(* IEC 61131-3 sources: 2026_Projet_YGO_ExcavatriceDragage/TOOLS/TEST_AUTO_CI/RESULTS/L_SIMULATION/tests (part 4) *)

(* ---- test_fb_simbench.st ---- *)
SETUP
VAR
    FB_Bench : FB_SimBench;
    FB_SimEnc : FB_Sim_Encoder;
    FB_SimJoy : FB_Sim_Joystick;
    FB_SimSafe : FB_Sim_Safety;
    FB_SimTrans : FB_Sim_Translation;
    RawPosM1 : UDINT := 0;
    RawPosM2 : UDINT := 0;
END_VAR
END_SETUP

TEST 'TC-P03-001 Dynamique Enable : neutralisation initiale, transition Ready au repos, puis coupure'
    (* Scan 0 : Enable=FALSE -> Neutralisation *)
    FB_Bench(Enable := FALSE, RawPosM1 := RawPosM1, RawPosM2 := RawPosM2);
    ASSERT_FALSE(FB_Bench.Ready, 'Enable=FALSE -> Ready=FALSE (neutralise)');

    ADVANCE_TIME(10000000);

    (* Scan 1 : Enable=TRUE -> SimBench actif *)
    FB_Bench(Enable := TRUE, RawPosM1 := RawPosM1, RawPosM2 := RawPosM2);
    ASSERT_TRUE(FB_Bench.Ready, 'Enable=TRUE -> Ready=TRUE (nominal)');

    ADVANCE_TIME(10000000);

    (* Scan 2 : Enable=FALSE -> Re-neutralisation *)
    FB_Bench(Enable := FALSE, RawPosM1 := RawPosM1, RawPosM2 := RawPosM2);
    ASSERT_FALSE(FB_Bench.Ready, 'Coupure -> Ready retombe a FALSE');
END_TEST

(* =========================================================================
   T419 — Reprise de jeu : ne jamais ouvrir la benne pendant une descente M1+M2.
   ========================================================================= *)

TEST 'TC-P13-074 T419 descente M1-M2 : compensation de fermeture conservee'
VAR
    CorrectionAfterAscentPts       : DINT;
    CorrectionAfterBothDescentPts  : DINT;
END_VAR
    (* La montee couplee etablit une compensation de fermeture observable. *)
    RawPosM1 := 1000000; RawPosM2 := 1100000;
    FB_Bench(Enable := TRUE, RawPosM1 := RawPosM1, RawPosM2 := RawPosM2,
             M1_RelayFwd := TRUE, M2_RelayFwd := TRUE,
             M1_BrakeCmd := TRUE, M2_BrakeCmd := TRUE,
             SimWinchCouplingModelActive := TRUE,
             M1_CablePos_M := 5.0, M2_CablePos_M := 18.5,
             BucketOffsetCloseM := 15.0, BucketCoherenceLimitM := 1.0);
    ADVANCE_TIME(10000000);

    (* Second scan : reprise de jeu de fermeture accumulee dans l'image M2. *)
    FB_Bench(Enable := TRUE, RawPosM1 := RawPosM1, RawPosM2 := RawPosM2,
             M1_RelayFwd := TRUE, M2_RelayFwd := TRUE,
             M1_BrakeCmd := TRUE, M2_BrakeCmd := TRUE,
             SimWinchCouplingModelActive := TRUE,
             M1_CablePos_M := 5.0, M2_CablePos_M := 18.5,
             BucketOffsetCloseM := 15.0, BucketCoherenceLimitM := 1.0);
    CorrectionAfterAscentPts := UDINT_TO_DINT(FB_Bench.Winch.COD2_PosValue) - UDINT_TO_DINT(RawPosM2);
    ASSERT_TRUE(CorrectionAfterAscentPts > 0, 'montee couplee -> compensation fermee presente');
    ADVANCE_TIME(10000000);

    (* Descente de charge M1+M2 : ce n'est pas une ouverture relative de la benne. *)
    FB_Bench(Enable := TRUE, RawPosM1 := RawPosM1, RawPosM2 := RawPosM2,
             M1_RelayFwd := FALSE, M1_RelayRev := TRUE,
             M2_RelayFwd := FALSE, M2_RelayRev := TRUE,
             M1_BrakeCmd := TRUE, M2_BrakeCmd := TRUE,
             SimWinchCouplingModelActive := TRUE,
             M1_CablePos_M := 5.0, M2_CablePos_M := 18.5,
             BucketOffsetCloseM := 15.0, BucketCoherenceLimitM := 1.0);
    CorrectionAfterBothDescentPts := UDINT_TO_DINT(FB_Bench.Winch.COD2_PosValue) - UDINT_TO_DINT(RawPosM2);
    ASSERT_EQ(CorrectionAfterBothDescentPts, CorrectionAfterAscentPts,
              'descente M1+M2 -> compensation de fermeture inchangee');
END_TEST

TEST 'TC-P13-075 T419 ouverture M2 seule : relachement borne conserve'
VAR
    CorrectionBeforeOpenPts : DINT;
    CorrectionAfterOpenPts  : DINT;
END_VAR
    (* Scenario autonome : etabli une fermeture avant l'ouverture relative M2 seule. *)
    RawPosM1 := 1000000; RawPosM2 := 1100000;
    FB_Bench(Enable := TRUE, RawPosM1 := RawPosM1, RawPosM2 := RawPosM2,
             M1_RelayFwd := TRUE, M2_RelayFwd := TRUE,
             M1_BrakeCmd := TRUE, M2_BrakeCmd := TRUE,
             SimWinchCouplingModelActive := TRUE,
             M1_CablePos_M := 5.0, M2_CablePos_M := 18.5,
             BucketOffsetCloseM := 15.0, BucketCoherenceLimitM := 1.0);
    ADVANCE_TIME(10000000);
    CorrectionBeforeOpenPts := UDINT_TO_DINT(FB_Bench.Winch.COD2_PosValue) - UDINT_TO_DINT(RawPosM2);
    ASSERT_TRUE(CorrectionBeforeOpenPts > 0, 'fermeture etablie avant ouverture M2 seule');
    ADVANCE_TIME(10000000);
    FB_Bench(Enable := TRUE, RawPosM1 := RawPosM1, RawPosM2 := RawPosM2,
             M1_RelayFwd := FALSE, M1_RelayRev := FALSE,
             M2_RelayFwd := FALSE, M2_RelayRev := TRUE,
             M2_BrakeCmd := TRUE,
             SimWinchCouplingModelActive := TRUE,
             M1_CablePos_M := 5.0, M2_CablePos_M := 18.5,
             BucketOffsetCloseM := 15.0, BucketCoherenceLimitM := 1.0);
    CorrectionAfterOpenPts := UDINT_TO_DINT(FB_Bench.Winch.COD2_PosValue) - UDINT_TO_DINT(RawPosM2);
    ASSERT_TRUE(CorrectionAfterOpenPts < CorrectionBeforeOpenPts,
                'ouverture M2 seule -> compensation relachee');
    ASSERT_TRUE((CorrectionBeforeOpenPts - CorrectionAfterOpenPts) <= 82,
                'ouverture M2 seule -> relachement borne a 0,02 m par scan');
END_TEST

TEST 'TC-P13-001 Sim_Safety : neutralisation sans Enable'
    FB_SimSafe(Enable := FALSE);
    ASSERT_FALSE(FB_SimSafe.SimChainOk, 'AU non ferme');
    ASSERT_FALSE(FB_SimSafe.SimContactorOk, 'Contacteur coupe');
END_TEST

(* =========================================================================
   AF-13 — FB_SimBench (TC-P13-010/011/012/013)
   ========================================================================= *)

TEST 'TC-P13-010 SimBench Enable=FALSE neutralise tout le banc'
    FB_Bench(Enable := FALSE, RawPosM1 := RawPosM1, RawPosM2 := RawPosM2);
    ASSERT_FALSE(FB_Bench.Ready, 'Enable=FALSE -> Ready=FALSE');
    ASSERT_FALSE(FB_Bench.Busy, 'Enable=FALSE -> Busy=FALSE');
    ASSERT_FALSE(FB_Bench.Done, 'Enable=FALSE -> Done=FALSE');
END_TEST

(* =========================================================================
   T342 — CR2 : reinjection silencieuse du comptage brut (RawPosM2 = 0 -> 1 100 000 pts)
   Remplace TC-P13-014 « initialise les codeurs absolus vierges » (ID par ailleurs porte
   par l'AF-13 pour le capteur haut TOP : collision d'ID levee au passage) : le banc
   n'initialise PLUS rien, le cas « memoire vierge » est couvert par l'initialisation
   declaree GVL_PERSISTENT._SimEncoderRawPosM1/M2 := 1000000.
   ========================================================================= *)

TEST 'TC-T342-010 AUCUNE reinjection du comptage brut : un 0 reel du codeur est conserve (pas de saut post-AU)'
    (* Etat EXACT de l'incident T338 (saut 8,50 -> 204,677 m apres reactivation du banc) :
       memoire codeur a 0, banc desactive (Enable=FALSE), puis reactivation du banc
       (GVL_Simulation.SimulationModeActive FALSE -> TRUE). Le comptage brut est un entier
       SIGNE dont le zero est arbitraire (correctif T338) : le banc ne doit JAMAIS y
       substituer une origine device, sous peine d'une teleportation de
       1 100 000 pts / 4096 pts/m = 268,55 m sur la position publiee, sans mouvement
       ni defaut, reference de homing conservee. *)
    FB_Bench(Enable := FALSE, RawPosM1 := RawPosM1, RawPosM2 := RawPosM2);
    RawPosM1 := 0;
    RawPosM2 := 0;
    ADVANCE_TIME(10000000);
    FB_Bench(Enable := TRUE, RawPosM1 := RawPosM1, RawPosM2 := RawPosM2);
    ASSERT_EQ(RawPosM2, 0, 'Reactivation : la memoire codeur M2 reste a 0 (aucune reinjection du banc)');
    ASSERT_EQ(FB_Bench.Winch.COD2_PosValue, 0, 'Aucun saut publie sur COD2_PosValue (268,55 m si reinjecte)');
    ASSERT_EQ(RawPosM1, 0, 'Reactivation : la memoire codeur M1 reste a 0 (aucune reinjection du banc)');
    ASSERT_EQ(FB_Bench.Winch.COD1_PosValue, 0, 'Aucun saut publie sur COD1_PosValue');
END_TEST

TEST 'TC-T342-011 Reactivation du banc : le comptage brut conserve sa valeur courante (aucune ecriture du banc)'
    (* Non-regression du meme invariant sur une memoire MID-COURSE (296 459 pts = la valeur
       R0 reconstituee par le diagnostic T338) : quelle que soit la valeur, la reactivation
       ne produit aucun ecart, et le banc reste sans ecriture sur la memoire du codeur. *)
    FB_Bench(Enable := FALSE, RawPosM1 := RawPosM1, RawPosM2 := RawPosM2);
    RawPosM1 := 296459;
    RawPosM2 := 296459;
    ADVANCE_TIME(10000000);
    FB_Bench(Enable := TRUE, RawPosM1 := RawPosM1, RawPosM2 := RawPosM2);
    ASSERT_EQ(RawPosM2, 296459, 'Memoire M2 mid-course inchangee par la reactivation du banc');
    ASSERT_EQ(FB_Bench.Winch.COD2_PosValue, 296459, 'Position publiee = comptage brut, sans ecart');
    ASSERT_EQ(RawPosM1, 296459, 'Memoire M1 mid-course inchangee par la reactivation du banc');
    ASSERT_EQ(FB_Bench.Winch.COD1_PosValue, 296459, 'Position publiee = comptage brut, sans ecart');
END_TEST

TEST 'TC-P13-011 SimBench 0 lecture GVL en interne (essai manuel — stub)'
    (* Stub : TC-P13-011 verifie que FB_SimBench ne lit aucune variable GVL_* en interne
       (toutes les entrees passees en parametres par PRG_02_Acquisition). Verification
       statique de code, non automatisable en boite noire. (essai manuel — stub) *)
    ASSERT_TRUE(TRUE, 'Stub : verification statique 0 lecture GVL (essai manuel)');
END_TEST

TEST 'TC-P13-012 SimBench polarite frein M1 : M1_BrakeIsOpen_DI := M1_BrakeCmd'
    FB_Bench(Enable := TRUE, M1_BrakeCmd := TRUE, RawPosM1 := RawPosM1, RawPosM2 := RawPosM2);
    ASSERT_TRUE(FB_Bench.Winch.M1_BrakeIsOpen_DI, 'M1_BrakeCmd=TRUE -> M1_BrakeIsOpen_DI=TRUE (jamais NOT)');
    ADVANCE_TIME(10000000);
    FB_Bench(Enable := TRUE, M1_BrakeCmd := FALSE, RawPosM1 := RawPosM1, RawPosM2 := RawPosM2);
    ASSERT_FALSE(FB_Bench.Winch.M1_BrakeIsOpen_DI, 'M1_BrakeCmd=FALSE -> M1_BrakeIsOpen_DI=FALSE');
END_TEST

TEST 'TC-T318-010 SimBench cable nominal independent du Kobold et injection explicite'
    FB_Bench(Enable := TRUE, SimKoboldContactValue := TRUE,
             SimM2TensionedCableFaultInject := FALSE,
             RawPosM1 := RawPosM1, RawPosM2 := RawPosM2);
    ASSERT_TRUE(FB_Bench.Winch.M2_TensionedCable_DI,
                'Kobold ne produit pas de mou de cable sans injection explicite');
    FB_Bench(Enable := TRUE, SimM2TensionedCableFaultInject := TRUE,
             RawPosM1 := RawPosM1, RawPosM2 := RawPosM2);
    ASSERT_FALSE(FB_Bench.Winch.M2_TensionedCable_DI,
                 'Injection explicite -> cable non tendu');
END_TEST

TEST 'TC-T318-020 Diagnostic electrique desactive publie etat neutre'
    FB_Bench(Enable := TRUE, SimWinchElectricalDiagnosticsActive := FALSE,
             RawPosM1 := RawPosM1, RawPosM2 := RawPosM2);
    ASSERT_EQ(FB_Bench.MotorTorqueM1_Nm, 0.0, 'Diagnostic M1 OFF -> couple neutre');
    ASSERT_FALSE(FB_Bench.MotorIsStalledM1, 'Diagnostic M1 OFF -> stall FALSE');
    ASSERT_EQ(FB_Bench.MotorTorqueM2_Nm, 0.0, 'Diagnostic M2 OFF -> couple neutre');
    ASSERT_FALSE(FB_Bench.MotorIsStalledM2, 'Diagnostic M2 OFF -> stall FALSE');
END_TEST

TEST 'TC-P13-015 SimBench delai frein M1 opt-in (T316) : SimWinchBrakeOpenDelayS retarde M1_BrakeIsOpen_DI sans jamais inverser la polarite'
    (* Delai desactive (0.0) : comportement historique, bascule au meme scan *)
    FB_Bench(Enable := TRUE, M1_BrakeCmd := TRUE, SimWinchBrakeOpenDelayS := 0.0, RawPosM1 := RawPosM1, RawPosM2 := RawPosM2);
    ASSERT_TRUE(FB_Bench.Winch.M1_BrakeIsOpen_DI, 'Delai=0.0 -> ouverture instantanee (non-regression)');
    ADVANCE_TIME(10000000);
    FB_Bench(Enable := TRUE, M1_BrakeCmd := FALSE, SimWinchBrakeOpenDelayS := 0.0, RawPosM1 := RawPosM1, RawPosM2 := RawPosM2);
    ASSERT_FALSE(FB_Bench.Winch.M1_BrakeIsOpen_DI, 'Retour delai=0.0 avant test delai>0 : etat repos');

    (* Delai actif (50 ms = 5 scans a 10 ms) : la DI reste fausse pendant le delai puis bascule *)
    ADVANCE_TIME(10000000);
    FB_Bench(Enable := TRUE, M1_BrakeCmd := TRUE, SimWinchDynamicsActive := TRUE, SimWinchBrakeOpenDelayS := 0.042, RawPosM1 := RawPosM1, RawPosM2 := RawPosM2);
    ASSERT_FALSE(FB_Bench.Winch.M1_BrakeIsOpen_DI, 'Scan 1/5 du delai : M1_BrakeIsOpen_DI reste FALSE, jamais TRUE en avance');
    ADVANCE_TIME(10000000);
    FB_Bench(Enable := TRUE, M1_BrakeCmd := TRUE, SimWinchDynamicsActive := TRUE, SimWinchBrakeOpenDelayS := 0.042, RawPosM1 := RawPosM1, RawPosM2 := RawPosM2);
    ASSERT_FALSE(FB_Bench.Winch.M1_BrakeIsOpen_DI, 'Scan 2/5 du delai : toujours FALSE');
    ADVANCE_TIME(10000000);
    FB_Bench(Enable := TRUE, M1_BrakeCmd := TRUE, SimWinchDynamicsActive := TRUE, SimWinchBrakeOpenDelayS := 0.042, RawPosM1 := RawPosM1, RawPosM2 := RawPosM2);
    ASSERT_FALSE(FB_Bench.Winch.M1_BrakeIsOpen_DI, 'Scan 3/5 du delai : toujours FALSE');
    ADVANCE_TIME(10000000);
    FB_Bench(Enable := TRUE, M1_BrakeCmd := TRUE, SimWinchDynamicsActive := TRUE, SimWinchBrakeOpenDelayS := 0.042, RawPosM1 := RawPosM1, RawPosM2 := RawPosM2);
    ASSERT_FALSE(FB_Bench.Winch.M1_BrakeIsOpen_DI, 'Scan 4/5 du delai : toujours FALSE');
    ADVANCE_TIME(10000000);
    FB_Bench(Enable := TRUE, M1_BrakeCmd := TRUE, SimWinchDynamicsActive := TRUE, SimWinchBrakeOpenDelayS := 0.042, RawPosM1 := RawPosM1, RawPosM2 := RawPosM2);
    ASSERT_TRUE(FB_Bench.Winch.M1_BrakeIsOpen_DI, 'Delai ecoule (5e scan) : M1_BrakeIsOpen_DI bascule TRUE');
END_TEST

TEST 'TC-T300-INT-010 SimBench M3 publie le retour dynamique du drive'
VAR
    i : INT;
END_VAR
    FB_Bench(Enable := TRUE, M3_ReqTremie := TRUE, M3_ReqMaintenance := FALSE,
             M3_SpeedCmd_Pct := 50.0, M3_BrakeCmd := TRUE,
             RawPosM1 := RawPosM1, RawPosM2 := RawPosM2);
    FOR i := 1 TO 20 DO
        FB_Bench(Enable := TRUE, M3_ReqTremie := TRUE, M3_ReqMaintenance := FALSE,
                 M3_SpeedCmd_Pct := 50.0, M3_BrakeCmd := TRUE,
                 RawPosM1 := RawPosM1, RawPosM2 := RawPosM2);
    END_FOR;
    ASSERT_EQ(FB_Bench.Translation.M3_StatusWord, 16#0087, 'M3 actif apres ouverture frein et retour frequence');
    FB_Bench(Enable := TRUE, M3_ReqTremie := FALSE, M3_ReqMaintenance := FALSE,
             M3_SpeedCmd_Pct := 0.0, M3_BrakeCmd := FALSE,
             RawPosM1 := RawPosM1, RawPosM2 := RawPosM2);
    FOR i := 1 TO 50 DO
        FB_Bench(Enable := TRUE, M3_ReqTremie := FALSE, M3_ReqMaintenance := FALSE,
                 M3_SpeedCmd_Pct := 0.0, M3_BrakeCmd := FALSE,
                 RawPosM1 := RawPosM1, RawPosM2 := RawPosM2);
    END_FOR;
    ASSERT_EQ(FB_Bench.Translation.M3_StatusWord, 16#0080, 'M3 arrete apres decroissance reelle de frequence');
END_TEST

TEST 'TC-T300-INT-030 Image SimBench relaye les DI M3 au decodeur production'
VAR
    Decoder : FB_Translation_PositionDecoder;
    HwInTranslation : ST_HwTranslation;
    i : INT;
END_VAR
    (* Le premier appel neutralise l'etat precedent. La copie explicite ci-dessous
       est representative du pont reel HwSim.Translation -> HwIn.Translation ;
       son unicite dans le programme est imposee statiquement par G502. *)
    FB_Bench(Enable := FALSE, RawPosM1 := RawPosM1, RawPosM2 := RawPosM2);
    FB_Bench(Enable := TRUE, M3_ReqTremie := FALSE, M3_ReqMaintenance := FALSE,
             M3_SpeedCmd_Pct := 0.0, M3_BrakeCmd := FALSE,
             RawPosM1 := RawPosM1, RawPosM2 := RawPosM2);
    HwInTranslation := FB_Bench.Translation;
    Decoder(SensorTremie := HwInTranslation.M3_PosTremie_DI,
            SensorPV := HwInTranslation.M3_PosPV_DI,
            SensorP2 := HwInTranslation.M3_PosPVP2_DI,
            SensorP1 := HwInTranslation.M3_PosP1_DI,
            SensorMaintenance := HwInTranslation.M3_PosMaintenance_DI);
    ASSERT_EQ(Decoder.SensorsWord, 2#00011, 'Repli P1 publie par l image puis decode sans injection aval');
    ASSERT_FALSE(Decoder.Incoherent, 'Mot P1 issu du SimBench coherent au decodeur production');

    (* T361 — 1800 scans (18 s) au lieu de 1100 : le banc a ete recale sur le gain odometrique
       reel (CST_M3FullTravelTimeS 8,0 -> 37,5 s, soit 0,8 m/s a 40 Hz au lieu de 3,75 m/s).
       Le trajet P1 (20 m) -> capteur Maintenance (29,95 m) demande desormais ~14 s
       (9,95 m a 0,8 m/s + ~2 s de rampe de frequence + ouverture du frein) : a 1100 scans le
       chariot n'atteignait plus la fin de course et le cas testait autre chose que son objet.
       Marge restante : ~4 s, soit ~3 m avant la butee mecanique. *)
    FOR i := 1 TO 1800 DO
        FB_Bench(Enable := TRUE, M3_ReqTremie := FALSE, M3_ReqMaintenance := TRUE,
                 M3_SpeedCmd_Pct := 100.0, M3_BrakeCmd := TRUE,
                 RawPosM1 := RawPosM1, RawPosM2 := RawPosM2);
        HwInTranslation := FB_Bench.Translation;
        Decoder(SensorTremie := HwInTranslation.M3_PosTremie_DI,
                SensorPV := HwInTranslation.M3_PosPV_DI,
                SensorP2 := HwInTranslation.M3_PosPVP2_DI,
                SensorP1 := HwInTranslation.M3_PosP1_DI,
                SensorMaintenance := HwInTranslation.M3_PosMaintenance_DI);
    END_FOR;
    ASSERT_EQ(Decoder.SensorsWord, 2#00000, 'Fin Maintenance dynamique traverse image et decodeur');
    ASSERT_TRUE(Decoder.LimitSwitchMaintenance, 'FDC Maintenance derive uniquement du mot image');
    ASSERT_FALSE(Decoder.Incoherent, 'Fin Maintenance dynamique reste coherente');
END_TEST

TEST 'TC-T300-INT-031 Intermittence P1 dynamique relayee au decodeur production'
VAR
    Decoder : FB_Translation_PositionDecoder;
    HwInTranslation : ST_HwTranslation;
    P1Previous : BOOL;
    P1Lost : BOOL := FALSE;
    P1Recovered : BOOL := FALSE;
    i : INT;
END_VAR
    FB_Bench(Enable := FALSE, RawPosM1 := RawPosM1, RawPosM2 := RawPosM2);
    FB_Bench(Enable := TRUE, M3_ReqTremie := FALSE, M3_ReqMaintenance := FALSE,
             M3_SpeedCmd_Pct := 0.0, M3_BrakeCmd := FALSE,
             RawPosM1 := RawPosM1, RawPosM2 := RawPosM2);
    HwInTranslation := FB_Bench.Translation;
    P1Previous := HwInTranslation.M3_PosP1_DI;

    (* Angle declencheur nul : l'episode est impose par la traversee mecanique,
       pas par un mot DI force. La graine et la periode restent deterministes. *)
    FOR i := 1 TO 1500 DO
        FB_Bench(Enable := TRUE, M3_ReqTremie := FALSE, M3_ReqMaintenance := TRUE,
                 M3_SpeedCmd_Pct := 100.0, M3_BrakeCmd := TRUE,
                 SimM3SensorIntermittenceActive := TRUE,
                 SimM3SensorStabilizationS := 1.0,
                 SimM3SensorIntermittencePeriodS := 0.12,
                 SimM3SensorElectricalDelayS := 0.0,
                 SimM3SensorLoadAngleTriggerRad := 0.0,
                 SimM3SensorScenarioSeed := 3001,
                 RawPosM1 := RawPosM1, RawPosM2 := RawPosM2);
        HwInTranslation := FB_Bench.Translation;
        Decoder(SensorTremie := HwInTranslation.M3_PosTremie_DI,
                SensorPV := HwInTranslation.M3_PosPV_DI,
                SensorP2 := HwInTranslation.M3_PosPVP2_DI,
                SensorP1 := HwInTranslation.M3_PosP1_DI,
                SensorMaintenance := HwInTranslation.M3_PosMaintenance_DI);
        IF P1Previous AND NOT HwInTranslation.M3_PosP1_DI THEN
            P1Lost := TRUE;
        END_IF;
        IF P1Lost AND HwInTranslation.M3_PosP1_DI THEN
            P1Recovered := TRUE;
        END_IF;
        P1Previous := HwInTranslation.M3_PosP1_DI;
    END_FOR;
    ASSERT_TRUE(P1Lost, 'P1 perd au moins une fois son etat pendant le franchissement');
    ASSERT_TRUE(P1Recovered, 'P1 est repris pendant l episode borne');
    ASSERT_FALSE(HwInTranslation.M3_PosP1_DI, 'P1 se stabilise a FALSE apres franchissement vers Maintenance');
    ASSERT_FALSE(Decoder.TranslationPosP1, 'Decodeur production voit la stabilisation du DI image');
END_TEST

TEST 'T196-003 Capteur haut manuel et polarite Free_DI correcte'
    FB_Bench(Enable := TRUE, SimTopPositionActive := TRUE,
             RawPosM1 := RawPosM1, RawPosM2 := RawPosM2);
    ASSERT_FALSE(FB_Bench.Winch.M1M2_TopPositionFree_DI,
                 'TopPositionActive=TRUE -> Free_DI=FALSE (capteur atteint)');
    ADVANCE_TIME(10000000);
    FB_Bench(Enable := TRUE, SimTopPositionActive := FALSE,
             RawPosM1 := RawPosM1, RawPosM2 := RawPosM2);
    ASSERT_TRUE(FB_Bench.Winch.M1M2_TopPositionFree_DI,
                'TopPositionActive=FALSE -> Free_DI=TRUE (butée libre)');
END_TEST

TEST 'T196-004 Capteur haut auto : forçage manuel SimTopPositionActive'
    FB_Bench(Enable := TRUE, SimTopPositionActive := FALSE,
             RawPosM1 := RawPosM1, RawPosM2 := RawPosM2);
    ASSERT_TRUE(FB_Bench.Winch.M1M2_TopPositionFree_DI,
                'SimTopPositionActive=FALSE -> capteur haut libre');
    ADVANCE_TIME(10000000);
    FB_Bench(Enable := TRUE, SimTopPositionActive := TRUE,
             RawPosM1 := RawPosM1, RawPosM2 := RawPosM2);
    ASSERT_FALSE(FB_Bench.Winch.M1M2_TopPositionFree_DI,
                 'SimTopPositionActive=TRUE -> capteur haut actif');
END_TEST

(* =========================================================================
   AF-13 — FB_Sim_Safety (TC-P13-020/021/022/023)
   ========================================================================= *)

TEST 'TC-P13-020 Sim_Safety SimChainOk = A AND B AND NOT BtnEmergencyStop'
    FB_SimSafe(Enable := TRUE, SimChainOkBit := TRUE, BtnEmergencyStop := FALSE);
    ADVANCE_TIME(60000000); (* Delai retombe relais 50ms *)
    FB_SimSafe(Enable := TRUE, SimChainOkBit := TRUE, BtnEmergencyStop := FALSE);
    ASSERT_TRUE(FB_SimSafe.SimChainOk, 'SimChainOkBit=TRUE -> SimChainOk=TRUE apres 50ms');

    ADVANCE_TIME(10000000);
    FB_SimSafe(Enable := TRUE, SimChainOkBit := FALSE, BtnEmergencyStop := FALSE);
    ADVANCE_TIME(60000000);
    FB_SimSafe(Enable := TRUE, SimChainOkBit := FALSE, BtnEmergencyStop := FALSE);
    ASSERT_FALSE(FB_SimSafe.SimChainOk, 'SimChainOkBit=FALSE -> SimChainOk=FALSE');

    ADVANCE_TIME(10000000);
    FB_SimSafe(Enable := TRUE, SimChainOkBit := TRUE, BtnEmergencyStop := TRUE);
    ADVANCE_TIME(60000000);
    FB_SimSafe(Enable := TRUE, SimChainOkBit := TRUE, BtnEmergencyStop := TRUE);
    ASSERT_FALSE(FB_SimSafe.SimChainOk, 'BtnEmergencyStop -> SimChainOk=FALSE');
END_TEST

TEST 'TC-P13-021 Sim_Safety SimContactorOk s auto-maintient sur EmergencyArming'
    FB_SimSafe(Enable := TRUE, SimChainOkBit := TRUE, EmergencyArming := FALSE, BtnEmergencyStop := FALSE);
    ADVANCE_TIME(60000000);
    FB_SimSafe(Enable := TRUE, SimChainOkBit := TRUE, EmergencyArming := FALSE, BtnEmergencyStop := FALSE);
    ASSERT_FALSE(FB_SimSafe.SimContactorOk, 'pas encore arme -> contacteur FALSE');

    (* Impulsion armement tenue 100ms *)
    ADVANCE_TIME(10000000);
    FB_SimSafe(Enable := TRUE, SimChainOkBit := TRUE, EmergencyArming := TRUE, BtnEmergencyStop := FALSE);
    ADVANCE_TIME(110000000);
    FB_SimSafe(Enable := TRUE, SimChainOkBit := TRUE, EmergencyArming := TRUE, BtnEmergencyStop := FALSE);
    ASSERT_TRUE(FB_SimSafe.SimContactorOk, 'EmergencyArming -> contacteur engage');

    (* Relachement impulsion -> auto-maintien *)
    ADVANCE_TIME(10000000);
    FB_SimSafe(Enable := TRUE, SimChainOkBit := TRUE, EmergencyArming := FALSE, BtnEmergencyStop := FALSE);
    ASSERT_TRUE(FB_SimSafe.SimContactorOk, 'auto-maintien : contacteur reste engage');

    (* Coupure chaine -> retombe apres chaine (50ms) + contacteur (50ms) *)
    ADVANCE_TIME(10000000);
    FB_SimSafe(Enable := TRUE, SimChainOkBit := FALSE, EmergencyArming := FALSE, BtnEmergencyStop := FALSE);
    ADVANCE_TIME(60000000); (* Chaine s ouvre *)
    FB_SimSafe(Enable := TRUE, SimChainOkBit := FALSE, EmergencyArming := FALSE, BtnEmergencyStop := FALSE);
    ADVANCE_TIME(60000000); (* Contacteur retombe *)
    FB_SimSafe(Enable := TRUE, SimChainOkBit := FALSE, EmergencyArming := FALSE, BtnEmergencyStop := FALSE);
    ASSERT_FALSE(FB_SimSafe.SimContactorOk, 'SimChainOk=FALSE -> contacteur retombe');
END_TEST

TEST 'TC-P13-022 Sim_Safety Enable=FALSE neutralise tout'
    FB_SimSafe(Enable := FALSE, PowerCutOff_A := TRUE, PowerCutOff_B := TRUE, EmergencyArming := TRUE, BtnEmergencyStop := FALSE);
    ASSERT_FALSE(FB_SimSafe.SimChainOk, 'Enable=FALSE -> SimChainOk=FALSE');
    ASSERT_FALSE(FB_SimSafe.SimContactorOk, 'Enable=FALSE -> SimContactorOk=FALSE');
END_TEST

TEST 'TC-P13-023 Sim_Safety latch AU non lie a la sim (essai manuel — stub)'
    (* Stub : TC-P13-023 verifie qu un defaut AU reel latche (RedundancyTestFailedCause /
       EmergencyArmingFailedCause dans FB_Safety_EmergencyManagementLogic) survit a la sim et
       ne se debloque que par front Reset runtime. Non automatisable en boite noire FB_Sim_Safety
       (latch dans le FB consommateur). (essai manuel — stub) *)
    ASSERT_TRUE(TRUE, 'Stub : latch AU a verifier manuellement (essai manuel)');
END_TEST

(* =========================================================================
   AF-13 — FB_Sim_Encoder (TC-P13-030/031/032/033)
   ========================================================================= *)

TEST 'TC-P13-030 Sim_Encoder RelayFwd/Rev font compter RawPos'
    RawPosM1 := 0;
    FB_SimEnc(Enable := TRUE, RelayFwd := TRUE, RelayRev := FALSE, StepNumber := 1, RawPos := RawPosM1);
    ASSERT_GT(FB_SimEnc.RawPosOut, 0, 'RelayFwd -> RawPos augmente');
    ADVANCE_TIME(10000000);
    RawPosM1 := 100;
    FB_SimEnc(Enable := TRUE, RelayFwd := TRUE, RelayRev := FALSE, StepNumber := 1, RawPos := RawPosM1);
    ASSERT_GT(FB_SimEnc.RawPosOut, 100, 'RelayFwd -> RawPos augmente depuis 100');
    ADVANCE_TIME(10000000);
    RawPosM1 := 100;
    FB_SimEnc(Enable := TRUE, RelayFwd := FALSE, RelayRev := TRUE, StepNumber := 1, RawPos := RawPosM1);
    ASSERT_LT(FB_SimEnc.RawPosOut, 100, 'RelayRev -> RawPos diminue');
END_TEST

TEST 'TC-P13-031 Sim_Encoder PresetCmd charge PresetValue'
    RawPosM1 := 0;
    FB_SimEnc(Enable := TRUE, RelayFwd := FALSE, RelayRev := FALSE, StepNumber := 1, PresetCmd := TRUE, PresetValue := 5000, RawPos := RawPosM1);
    ADVANCE_TIME(10000000);
    FB_SimEnc(Enable := TRUE, RelayFwd := FALSE, RelayRev := FALSE, StepNumber := 1, PresetCmd := FALSE, PresetValue := 5000, RawPos := RawPosM1);
    ADVANCE_TIME(10000000);
    FB_SimEnc(Enable := TRUE, RelayFwd := FALSE, RelayRev := FALSE, StepNumber := 1, PresetCmd := FALSE, PresetValue := 5000, RawPos := RawPosM1);
    ADVANCE_TIME(10000000);
    FB_SimEnc(Enable := TRUE, RelayFwd := FALSE, RelayRev := FALSE, StepNumber := 1, PresetCmd := FALSE, PresetValue := 5000, RawPos := RawPosM1);
    ASSERT_EQ(FB_SimEnc.RawPosOut, 5000, 'Preset applique apres latence');
END_TEST

TEST 'TC-P13-032 Sim_Encoder le comptage franchit 0 au lieu de s y figer (butee silencieuse supprimee, T338)'
    (* Realigne sur la semantique T338 (comptage brut SIGNED 32 bits) : cette copie etait restee
       sur l'ancienne butee `RawPos := 0`, ce qui rendait la suite FB_SimBench ROUGE (41/42) sur
       HEAD depuis le commit 6a5910da — non-regression T338 incomplete. *)
    RawPosM1 := 41; (* 41 pts = exactement un pas de descente au palier 1 (1,0 x 4096 x 0,010) *)
    FB_SimEnc(Enable := TRUE, RelayFwd := FALSE, RelayRev := TRUE, StepNumber := 1, RawPos := RawPosM1);
    RawPosM1 := FB_SimEnc.RawPosOut; (* le caller conserve la memoire persistante du codeur *)
    ASSERT_EQ(FB_SimEnc.RawPosOut, 0, 'Un pas de descente amene le comptage exactement a 0 (point de passage)');
    ADVANCE_TIME(10000000);
    FB_SimEnc(Enable := TRUE, RelayFwd := FALSE, RelayRev := TRUE, StepNumber := 1, RawPos := RawPosM1);
    RawPosM1 := FB_SimEnc.RawPosOut;
    ASSERT_TRUE(FB_SimEnc.RawPosOut <> 0, 'Scan suivant : le comptage franchit 0 au lieu de s y figer');
    ASSERT_EQ(FB_SimEnc.RawPosOut, 4294967255, 'Comptage = -41 pts (aucune borne a 0, 2^32 - 41 en signe)');
END_TEST

TEST 'TC-P13-033 Sim_Encoder RawPos survit a un reset froid (essai manuel — stub)'
    (* Stub : TC-P13-033 verifie que RawPos (VAR_IN_OUT reference GVL_PERSISTENT) survit a un
       reset froid. Non automatisable en boite noire (depend de la persistance CODESYS).
       (essai manuel — stub) *)
    ASSERT_TRUE(TRUE, 'Stub : persistance RawPos a verifier manuellement (essai manuel)');
END_TEST

(* =========================================================================
   AF-13 — FB_Sim_Translation (TC-P13-040/041/042/043)
   ========================================================================= *)

TEST 'TC-T300-INT-020 Sim_Translation initialise le mot P1'
    FB_SimTrans(Enable := TRUE, ReqTremie := FALSE, ReqMaintenance := FALSE,
                SpeedTgt_Pct := 0.0, BrakeReleaseCmd := FALSE);
    ASSERT_FALSE(FB_SimTrans.PosTremie, 'P1 ne doit pas annoncer Tremie');
    ASSERT_FALSE(FB_SimTrans.PosPV, 'P1 ne doit pas annoncer PV');
    ASSERT_FALSE(FB_SimTrans.PosP2, 'P1 ne doit pas annoncer P2');
    ASSERT_TRUE(FB_SimTrans.PosP1, 'P1 actif au repli');
    ASSERT_TRUE(FB_SimTrans.PosMaintenance, 'Mot thermometre P1 coherent');
END_TEST

TEST 'TC-T300-INT-021 Sim_Translation neutralise deux sens simultanes'
    FB_SimTrans(Enable := TRUE, ReqTremie := TRUE, ReqMaintenance := TRUE,
                SpeedTgt_Pct := 100.0, BrakeReleaseCmd := TRUE);
    ASSERT_EQ(FB_SimTrans.FrequencyCmd_Hz, 0.0, 'Deux sens ne creent aucune consigne');
    ASSERT_EQ(FB_SimTrans.ActualFrequency_Hz, 0.0, 'Aucun retour variateur sans sens unique');
END_TEST

TEST 'TC-T300-INT-022 Sim_Translation borne et publie la fin de course Maintenance'
VAR
    i : INT;
END_VAR
    FB_SimTrans(Enable := FALSE);
    FB_SimTrans(Enable := TRUE, ReqTremie := FALSE, ReqMaintenance := TRUE,
                SpeedTgt_Pct := 100.0, FullTravelTimeS := 0.5,
                BrakeReleaseCmd := TRUE, SensorElectricalDelayS := 0.0);
    FOR i := 1 TO 400 DO
        FB_SimTrans(Enable := TRUE, ReqTremie := FALSE, ReqMaintenance := TRUE,
                    SpeedTgt_Pct := 100.0, FullTravelTimeS := 0.5,
                    BrakeReleaseCmd := TRUE, SensorElectricalDelayS := 0.0);
    END_FOR;
    ASSERT_GE(FB_SimTrans.PositionTrue_M, 0.0, 'Borne Tremie respectee');
    ASSERT_LE(FB_SimTrans.PositionTrue_M, 30.0, 'Borne Maintenance respectee');
    ASSERT_FALSE(FB_SimTrans.PosMaintenance, 'Maintenance publie le mot 00000 a la butee');
END_TEST

TEST 'TC-T300-INT-023 Sim_Translation desactive se replie P1'
    FB_SimTrans(Enable := FALSE, ReqTremie := FALSE, ReqMaintenance := TRUE,
                SpeedTgt_Pct := 100.0, BrakeReleaseCmd := TRUE);
    ASSERT_EQ(FB_SimTrans.PositionTrue_M, 20.0, 'Repli physique P1');
    ASSERT_TRUE(FB_SimTrans.PosP1, 'Capteur P1 coherent hors simulation');
    ASSERT_TRUE(FB_SimTrans.PosMaintenance, 'Mot P1 coherent hors simulation');
    ASSERT_FALSE(FB_SimTrans.BrakeContactOpen, 'Frein confirme ferme hors simulation');
END_TEST

(* =========================================================================
   AF-13 — FB_Sim_Joystick (TC-P13-050/051/052)
   ========================================================================= *)

TEST 'TC-P13-050 Sim_Joystick initialise au neutre au premier cycle'
    FB_SimJoy(Enable := TRUE, NeutralRaw := 5000, MaxRaw := 10000);
    ASSERT_EQ(FB_SimJoy.RawX, 5000, 'premier cycle -> RawX=NeutralRaw');
    ASSERT_EQ(FB_SimJoy.RawY, 5000, 'premier cycle -> RawY=NeutralRaw');
    ASSERT_FALSE(FB_SimJoy.RawButton, 'premier cycle -> RawButton=FALSE');
END_TEST

TEST 'TC-P13-051 Sim_Joystick sorties forçables en instance (essai manuel — stub)'
    (* Stub : TC-P13-051 verifie que RawX/RawY/RawButton restent forçables librement en instance
       CODESYS apres l'init (le FB n'ecrit plus ces sorties apres le premier cycle). Non
       automatisable en boite noire (depend du forçage CODESYS). (essai manuel — stub) *)
    ASSERT_TRUE(TRUE, 'Stub : forçage joystick a verifier manuellement (essai manuel)');
END_TEST

TEST 'TC-P13-052 Sim_Joystick homme-mort : RawButton reflete l appui (partie AUTO)'
    (* Aucun bouton -> RawButton=FALSE *)
    FB_SimJoy(Enable := TRUE, NeutralRaw := 5000, MaxRaw := 10000);
    ASSERT_FALSE(FB_SimJoy.RawButton, 'aucun bouton -> RawButton=FALSE');
    ADVANCE_TIME(10000000);
    (* Bouton directionnel actif -> RawButton=TRUE (homme-mort inclus) *)
    FB_SimJoy(Enable := TRUE, NeutralRaw := 5000, MaxRaw := 10000, BtnRight_Fwd_MAINT := TRUE);
    ASSERT_TRUE(FB_SimJoy.RawButton, 'bouton actif -> RawButton=TRUE');
END_TEST

(* =========================================================================
   AF-13 — FB_SimBench : rattrapage mecanique M1/M2 (T328)
   Plan : DOC/WFLOW/CONTRACTS/PLAN_T328_SIMBENCH_COUPLAGE_MECANIQUE_M1M2.md
   ========================================================================= *)

TEST 'TC-P13-060 T328 montee couplee : rattrapage actif et correction bornee'
    (* Montée couplée réelle (relais M1+M2 même sens, freins desserrés), benne DANS le trou métier
       T327 : écart 13,5 m < entrée de bande fermée (14,5 m). Le rattrapage agit, borné par la pente. *)
    RawPosM1 := 1000000; RawPosM2 := 1100000;
    FB_Bench(Enable := TRUE, RawPosM1 := RawPosM1, RawPosM2 := RawPosM2,
             M1_RelayFwd := TRUE, M2_RelayFwd := TRUE,
             M1_BrakeCmd := TRUE, M2_BrakeCmd := TRUE,
             SimWinchCouplingModelActive := TRUE,
             M1_CablePos_M := 5.0, M2_CablePos_M := 18.5,
             BucketOffsetCloseM := 15.0, BucketCoherenceLimitM := 1.0);
    ASSERT_TRUE(FB_Bench.WinchCouplingActive, 'montee couplee -> rattrapage actif');
    ASSERT_TRUE(FB_Bench.WinchCouplingCorrectionPts > 0, 'ecart sous la bande -> correction non nulle');
    ASSERT_TRUE(FB_Bench.WinchCouplingCorrectionPts <= 82, 'correction bornee (0,02 m/scan = 82 points)');
    ASSERT_TRUE(FB_Bench.Winch.COD2_PosValue > RawPosM2, 'correction appliquee a l IMAGE M2 uniquement');
END_TEST

TEST 'TC-P13-061 T328 arret et jog M2 seul : ecart fige, aucune correction'
    (* Relais à 0 : aucun mouvement réel -> jamais de rattrapage (AC6). *)
    FB_Bench(Enable := TRUE, RawPosM1 := RawPosM1, RawPosM2 := RawPosM2,
             M1_RelayFwd := FALSE, M2_RelayFwd := FALSE,
             SimWinchCouplingModelActive := TRUE,
             M1_CablePos_M := 5.0, M2_CablePos_M := 18.5,
             BucketOffsetCloseM := 15.0, BucketCoherenceLimitM := 1.0);
    ASSERT_FALSE(FB_Bench.WinchCouplingActive, 'relais a 0 -> pas de rattrapage');
    ASSERT_EQ(FB_Bench.WinchCouplingCorrectionPts, 0, 'aucune correction a l arret');
    ASSERT_EQ(FB_Bench.Winch.COD2_PosValue, RawPosM2, 'image M2 inchangee a l arret');
    ADVANCE_TIME(10000000);
    (* Jog M2 seul (un seul treuil actif) -> toujours aucun rattrapage *)
    FB_Bench(Enable := TRUE, RawPosM1 := RawPosM1, RawPosM2 := RawPosM2,
             M1_RelayFwd := FALSE, M2_RelayFwd := TRUE,
             M1_BrakeCmd := FALSE, M2_BrakeCmd := TRUE,
             SimWinchCouplingModelActive := TRUE,
             M1_CablePos_M := 5.0, M2_CablePos_M := 18.5,
             BucketOffsetCloseM := 15.0, BucketCoherenceLimitM := 1.0);
    ASSERT_FALSE(FB_Bench.WinchCouplingActive, 'jog M2 seul -> pas de rattrapage');
    ASSERT_EQ(FB_Bench.WinchCouplingCorrectionPts, 0, 'jog M2 seul -> aucune correction');
END_TEST

TEST 'TC-P13-062 T328 machoires bloquees : rattrapage inhibe et charge forcee'
    FB_Bench(Enable := TRUE, RawPosM1 := RawPosM1, RawPosM2 := RawPosM2,
             M1_RelayFwd := TRUE, M2_RelayFwd := TRUE,
             M1_BrakeCmd := TRUE, M2_BrakeCmd := TRUE,
             SimWinchCouplingModelActive := TRUE,
             SimBucketJamActive := TRUE,
             SimWinchElectricalDiagnosticsActive := TRUE,
             M1_CablePos_M := 5.0, M2_CablePos_M := 18.5,
             BucketOffsetCloseM := 15.0, BucketCoherenceLimitM := 1.0);
    ASSERT_FALSE(FB_Bench.WinchCouplingActive, 'blocage machoires -> rattrapage inhibe');
    ASSERT_EQ(FB_Bench.WinchCouplingCorrectionPts, 0, 'blocage -> aucune correction');
    ASSERT_TRUE(FB_Bench.MotorTorqueM1_Nm > 0.0, 'blocage -> charge forcee observable (diagnostic)');
END_TEST

TEST 'TC-P13-063 T328 modele desactive : image M2 inchangee (non-masquage T327)'
    FB_Bench(Enable := TRUE, RawPosM1 := RawPosM1, RawPosM2 := RawPosM2,
             M1_RelayFwd := TRUE, M2_RelayFwd := TRUE,
             M1_BrakeCmd := TRUE, M2_BrakeCmd := TRUE,
             SimWinchCouplingModelActive := FALSE,
             M1_CablePos_M := 5.0, M2_CablePos_M := 18.5,
             BucketOffsetCloseM := 15.0, BucketCoherenceLimitM := 1.0);
    ASSERT_FALSE(FB_Bench.WinchCouplingActive, 'modele OFF -> pas de rattrapage');
    ASSERT_EQ(FB_Bench.WinchCouplingCorrectionPts, 0, 'modele OFF -> aucune correction');
    ASSERT_EQ(FB_Bench.Winch.COD2_PosValue, RawPosM2, 'modele OFF -> image M2 identique (trou T327 preserve)');
END_TEST

TEST 'TC-P13-064 T328 cable mou : rattrapage inhibe (aucun effort transmis)'
    FB_Bench(Enable := TRUE, RawPosM1 := RawPosM1, RawPosM2 := RawPosM2,
             M1_RelayFwd := TRUE, M2_RelayFwd := TRUE,
             M1_BrakeCmd := TRUE, M2_BrakeCmd := TRUE,
             SimWinchCouplingModelActive := TRUE,
             SimM2TensionedCableFaultInject := TRUE,
             M1_CablePos_M := 5.0, M2_CablePos_M := 18.5,
             BucketOffsetCloseM := 15.0, BucketCoherenceLimitM := 1.0);
    ASSERT_FALSE(FB_Bench.WinchCouplingActive, 'cable mou -> pas de rattrapage');
END_TEST

TEST 'TC-P13-065 T328 banc eteint : image reelle repliquee sans correction'
    FB_Bench(Enable := FALSE, RawPosM1 := RawPosM1, RawPosM2 := RawPosM2,
             M1_RelayFwd := TRUE, M2_RelayFwd := TRUE,
             M1_BrakeCmd := TRUE, M2_BrakeCmd := TRUE,
             SimWinchCouplingModelActive := TRUE,
             M1_CablePos_M := 5.0, M2_CablePos_M := 18.5,
             BucketOffsetCloseM := 15.0, BucketCoherenceLimitM := 1.0);
    ASSERT_FALSE(FB_Bench.WinchCouplingActive, 'banc desactive -> aucun rattrapage');
    ASSERT_EQ(FB_Bench.Winch.COD2_PosValue, RawPosM2, 'banc desactive -> image sans correction');
END_TEST

TEST 'TC-P13-066 T328 convergence multi-scan du rattrapage vers la bande fermee'
VAR
    i        : INT;
    M2_Pos_M : REAL := 0.0;
END_VAR
    (* Boucle fermee simulee : la position M2 vue par le metier suit l'image corrigee, comme dans la
       chaine reelle (HwSim -> HwIn -> codeur). Delta initial 13,5 m = trou metier de fermeture.
       Chaque appel du FB vaut un scan de 10 ms (le modele utilise CST_SimBenchCycleTimeS, pas le
       temps du harness) : la boucle n'avance donc pas le temps du harness. *)
    RawPosM1 := 1000000; RawPosM2 := 1100000;
    M2_Pos_M := 18.5;   (* Delta = M2 - M1 = 13,5 m *)
    FOR i := 1 TO 100 DO
        FB_Bench(Enable := TRUE, RawPosM1 := RawPosM1, RawPosM2 := RawPosM2,
                 M1_RelayFwd := TRUE, M2_RelayFwd := TRUE,
                 M1_BrakeCmd := TRUE, M2_BrakeCmd := TRUE,
                 SimWinchCouplingModelActive := TRUE,
                 M1_CablePos_M := 5.0, M2_CablePos_M := M2_Pos_M,
                 BucketOffsetCloseM := 15.0, BucketCoherenceLimitM := 1.0);
        ASSERT_TRUE(FB_Bench.WinchCouplingCorrectionPts <= 82, 'correction bornee a 0,02 m par scan');
        M2_Pos_M := M2_Pos_M + DINT_TO_REAL(FB_Bench.WinchCouplingCorrectionPts) * (2.0 / 8192.0);
    END_FOR;
    ADVANCE_TIME(10000000);
    ASSERT_TRUE((M2_Pos_M - 5.0) >= 14.0, 'Delta entre dans la bande fermee (>= 14,0 m) en temps borne');
END_TEST

TEST 'TC-P13-067 T328 un preset purge l offset de reprise de jeu (image = codeur)'
    RawPosM1 := 1000000; RawPosM2 := 1100000;
    (* Session active : un offset est bien accumule. *)
    FB_Bench(Enable := TRUE, RawPosM1 := RawPosM1, RawPosM2 := RawPosM2,
             M1_RelayFwd := TRUE, M2_RelayFwd := TRUE,
             M1_BrakeCmd := TRUE, M2_BrakeCmd := TRUE,
             SimWinchCouplingModelActive := TRUE,
             M1_CablePos_M := 5.0, M2_CablePos_M := 18.5,
             BucketOffsetCloseM := 15.0, BucketCoherenceLimitM := 1.0);
    ASSERT_TRUE(FB_Bench.Winch.COD2_PosValue > RawPosM2, 'offset de reprise de jeu accumule');
    ADVANCE_TIME(10000000);
    (* Preset M2 (PresetTriggerCmd = 2) : la reference absolue est reecrite -> offset purge. *)
    FB_Bench(Enable := TRUE, RawPosM1 := RawPosM1, RawPosM2 := RawPosM2,
             M1_RelayFwd := TRUE, M2_RelayFwd := TRUE,
             M1_BrakeCmd := TRUE, M2_BrakeCmd := TRUE,
             SimWinchCouplingModelActive := TRUE, M2_PresetTriggerCmd := 2,
             M1_CablePos_M := 5.0, M2_CablePos_M := 18.5,
             BucketOffsetCloseM := 15.0, BucketCoherenceLimitM := 1.0);
    ASSERT_EQ(FB_Bench.Winch.COD2_PosValue, RawPosM2, 'preset -> offset purge, image = codeur');
END_TEST

TEST 'TC-P13-068 T328 mode OFF apres session active : aucun offset residuel'
    RawPosM1 := 1000000; RawPosM2 := 1100000;
    FB_Bench(Enable := TRUE, RawPosM1 := RawPosM1, RawPosM2 := RawPosM2,
             M1_RelayFwd := TRUE, M2_RelayFwd := TRUE,
             M1_BrakeCmd := TRUE, M2_BrakeCmd := TRUE,
             SimWinchCouplingModelActive := TRUE,
             M1_CablePos_M := 5.0, M2_CablePos_M := 18.5,
             BucketOffsetCloseM := 15.0, BucketCoherenceLimitM := 1.0);
    ASSERT_TRUE(FB_Bench.Winch.COD2_PosValue > RawPosM2, 'offset accumule en mode actif');
    ADVANCE_TIME(10000000);
    (* Bascule mode OFF : l'image doit redevenir strictement celle du codeur (non-masquage). *)
    FB_Bench(Enable := TRUE, RawPosM1 := RawPosM1, RawPosM2 := RawPosM2,
             M1_RelayFwd := TRUE, M2_RelayFwd := TRUE,
             M1_BrakeCmd := TRUE, M2_BrakeCmd := TRUE,
             SimWinchCouplingModelActive := FALSE,
             M1_CablePos_M := 5.0, M2_CablePos_M := 18.5,
             BucketOffsetCloseM := 15.0, BucketCoherenceLimitM := 1.0);
    ASSERT_FALSE(FB_Bench.WinchCouplingActive, 'mode OFF -> rattrapage inactif');
    ASSERT_EQ(FB_Bench.Winch.COD2_PosValue, RawPosM2, 'mode OFF -> aucun offset residuel sur l image');
END_TEST

(* =========================================================================
   T328 (reprise DSH03) — SCENARIO UTILISATEUR 2026-09-20 : benne FERMEE avec
   ecart residuel ~5 % (voyant ferme allume), puis MONTEE couplee.
   Definitions (source FB_Bucket.st:591 + GVL_PERSISTENT.st:66-70) :
     Ouverture_Pct = 100 * (OffsetCloseM - Delta) / (OffsetCloseM - OffsetOpenM)
     Delta = CablePosM2 - CablePosM1 ; OffsetCloseM = 15,0 m ; OffsetOpenM = 0,0 m
     => ecart 5 %  <=> Delta = 14,25 m   (=> IsClosed TRUE : Delta >= 14,0 m)
        ecart 0 %  <=> Delta = 15,0 m   (butee mecanique benne fermee)
        ecart 3,33 % <=> Delta = 14,50 m (cible ABANDONNEE (plafonnait l ecart a 3,4 %), FB_SimBench.st:505)
   Aucun de ces cas n existait dans la suite : TC-P13-060..068 partent tous de
   Delta = 13,5 m (10 % ouverture, trou metier T327), jamais du residuel POST-fermeture.
   CIBLE RETENUE (arbitrage CC01 2026-09-20, D1) : BUTEE mecanique (ecart 0 %).
   ========================================================================= *)

TEST 'TC-P13-070 T328 scenario utilisateur : ecart 5 % (Delta 14,25 m) resorbe vers 0 % en montee couplee'
VAR
    i        : INT;
    M2_Pos_M : REAL := 0.0;
END_VAR
    (* Boucle fermee reelle : HwSim (image corrigee) -> HwIn -> codeur M2 -> Delta mesure. *)
    RawPosM1 := 1000000; RawPosM2 := 1100000;
    M2_Pos_M := 14.25 + 5.0;   (* Delta initial = 14,25 m => ouverture 5 % (cas utilisateur) *)
    FOR i := 1 TO 800 DO
        FB_Bench(Enable := TRUE, RawPosM1 := RawPosM1, RawPosM2 := RawPosM2,
                 M1_RelayFwd := TRUE, M2_RelayFwd := TRUE,
                 M1_BrakeCmd := TRUE, M2_BrakeCmd := TRUE,
                 SimWinchCouplingModelActive := TRUE,
                 M1_CablePos_M := 5.0, M2_CablePos_M := M2_Pos_M,
                 BucketOffsetCloseM := 15.0, BucketCoherenceLimitM := 1.0);
        ASSERT_TRUE(FB_Bench.WinchCouplingCorrectionPts <= 82, 'correction bornee a 0,02 m par scan');
        M2_Pos_M := M2_Pos_M + DINT_TO_REAL(FB_Bench.WinchCouplingCorrectionPts) * (2.0 / 8192.0);
    END_FOR;
    ADVANCE_TIME(10000000);
    (* Plancher de quantification : arret des que l increment < 1 point codeur (0,244 mm)
       => ecart residuel <= 2,5 cm soit 0,17 %, affiche 0 % a l IHM. *)
    ASSERT_TRUE((M2_Pos_M - 5.0) >= 14.97, 'ECART ATTENDU 0 % (Delta -> butee 15,0 m) pendant la montee');
    ASSERT_TRUE((M2_Pos_M - 5.0) <= 15.0, 'jamais de depassement de la butee mecanique');
END_TEST

TEST 'TC-P13-071 T328 cible : le point fixe du modele EST la butee mecanique (ecart 0 %)'
VAR
    i        : INT;
    M2_Pos_M : REAL := 0.0;
END_VAR
    (* Meme scenario que TC-P13-070 : on MESURE le point fixe du modele apres correctif D1.
       Cible = OffsetCloseM = 15,00 m ; point fixe mesure >= 14,975 m : le modele s arrete des que
       l increment 1er ordre devient < 1 point codeur (0,244 mm), soit un residu <= 2,5 cm.
       => ouverture residuelle <= 0,17 %, jamais un plancher de 3,4 %. *)
    RawPosM1 := 1000000; RawPosM2 := 1100000;
    M2_Pos_M := 14.25 + 5.0;
    FOR i := 1 TO 800 DO
        FB_Bench(Enable := TRUE, RawPosM1 := RawPosM1, RawPosM2 := RawPosM2,
                 M1_RelayFwd := TRUE, M2_RelayFwd := TRUE,
                 M1_BrakeCmd := TRUE, M2_BrakeCmd := TRUE,
                 SimWinchCouplingModelActive := TRUE,
                 M1_CablePos_M := 5.0, M2_CablePos_M := M2_Pos_M,
                 BucketOffsetCloseM := 15.0, BucketCoherenceLimitM := 1.0);
        M2_Pos_M := M2_Pos_M + DINT_TO_REAL(FB_Bench.WinchCouplingCorrectionPts) * (2.0 / 8192.0);
    END_FOR;
    ADVANCE_TIME(10000000);
    ASSERT_NEAR(M2_Pos_M - 5.0, 15.0, 0.03);
    ASSERT_TRUE((M2_Pos_M - 5.0) <= 15.0, 'point fixe = butee, jamais au-dela');
END_TEST

TEST 'TC-P13-072 T328 sur-fermeture (Delta > butee) : ecart FIGE, jamais corrige'
VAR
    i        : INT;
    M2_Pos_M : REAL := 0.0;
END_VAR
    (* Decision CC01 2026-09-20 (D2) : une sur-fermeture (Delta 15,75 m, soit +5 % AU-DELA de la
       butee 15,0 m, toujours dans la bande fermee 14,0..16,0 m) n est PAS corrigee : le modele
       reste strictement unidirectionnel -> rouvrir la benne pour resorber une sur-fermeture
       serait un mouvement non commande. Ecart FIGE : comportement voulu et teste. *)
    RawPosM1 := 1000000; RawPosM2 := 1100000;
    M2_Pos_M := 15.75 + 5.0;
    FOR i := 1 TO 100 DO
        FB_Bench(Enable := TRUE, RawPosM1 := RawPosM1, RawPosM2 := RawPosM2,
                 M1_RelayFwd := TRUE, M2_RelayFwd := TRUE,
                 M1_BrakeCmd := TRUE, M2_BrakeCmd := TRUE,
                 SimWinchCouplingModelActive := TRUE,
                 M1_CablePos_M := 5.0, M2_CablePos_M := M2_Pos_M,
                 BucketOffsetCloseM := 15.0, BucketCoherenceLimitM := 1.0);
        ASSERT_EQ(FB_Bench.WinchCouplingCorrectionPts, 0, 'sur-fermeture 5 % -> aucune correction');
        M2_Pos_M := M2_Pos_M + DINT_TO_REAL(FB_Bench.WinchCouplingCorrectionPts) * (2.0 / 8192.0);
    END_FOR;
    ADVANCE_TIME(10000000);
    ASSERT_NEAR(M2_Pos_M - 5.0, 15.75, 0.01);
END_TEST

TEST 'TC-P13-073 T328 GARDE-FOU : toute la bande de residus post-fermeture converge vers la butee'
VAR
    i        : INT;
    M2_Pos_M : REAL := 0.0;
END_VAR
    (* Garde-fou du trou de test qui a laisse passer T328 : la suite livree ne testait QUE
       Delta = 13,5 m. On couvre la bande des residus POST-fermeture reellement produite par la
       coupure d'anticipation + le roulis : 13,8 m (coupure T327) / 14,25 m (cas utilisateur 5 %) /
       14,75 m (haut de bande). Les trois doivent rejoindre la butee (ecart 0 %).
       (3 scenarios deroules : le harnais n accepte pas les boucles FOR imbriquees.) *)
    RawPosM1 := 1000000; RawPosM2 := 1100000;

    (* --- Residu 13,8 m (coupure d'anticipation T327) --- *)
    M2_Pos_M := 13.8 + 5.0;
    FOR i := 1 TO 800 DO
        FB_Bench(Enable := TRUE, RawPosM1 := RawPosM1, RawPosM2 := RawPosM2,
                 M1_RelayFwd := TRUE, M2_RelayFwd := TRUE,
                 M1_BrakeCmd := TRUE, M2_BrakeCmd := TRUE,
                 SimWinchCouplingModelActive := TRUE,
                 M1_CablePos_M := 5.0, M2_CablePos_M := M2_Pos_M,
                 BucketOffsetCloseM := 15.0, BucketCoherenceLimitM := 1.0);
        ASSERT_TRUE(FB_Bench.WinchCouplingCorrectionPts <= 82, 'correction bornee a 0,02 m par scan');
        M2_Pos_M := M2_Pos_M + DINT_TO_REAL(FB_Bench.WinchCouplingCorrectionPts) * (2.0 / 8192.0);
    END_FOR;
    ADVANCE_TIME(10000000);
    ASSERT_TRUE((M2_Pos_M - 5.0) >= 14.97, 'residu 13,8 m -> butee atteinte (ecart <= 0,2 %)');
    ASSERT_TRUE((M2_Pos_M - 5.0) <= 15.0, 'residu 13,8 m -> aucun depassement de butee');

    (* --- Residu 14,25 m (cas utilisateur : ecart 5 %, voyant ferme allume) --- *)
    M2_Pos_M := 14.25 + 5.0;
    FOR i := 1 TO 800 DO
        FB_Bench(Enable := TRUE, RawPosM1 := RawPosM1, RawPosM2 := RawPosM2,
                 M1_RelayFwd := TRUE, M2_RelayFwd := TRUE,
                 M1_BrakeCmd := TRUE, M2_BrakeCmd := TRUE,
                 SimWinchCouplingModelActive := TRUE,
                 M1_CablePos_M := 5.0, M2_CablePos_M := M2_Pos_M,
                 BucketOffsetCloseM := 15.0, BucketCoherenceLimitM := 1.0);
        ASSERT_TRUE(FB_Bench.WinchCouplingCorrectionPts <= 82, 'correction bornee a 0,02 m par scan');
        M2_Pos_M := M2_Pos_M + DINT_TO_REAL(FB_Bench.WinchCouplingCorrectionPts) * (2.0 / 8192.0);
    END_FOR;
    ADVANCE_TIME(10000000);
    ASSERT_TRUE((M2_Pos_M - 5.0) >= 14.97, 'residu 14,25 m -> butee atteinte (ecart <= 0,2 %)');
    ASSERT_TRUE((M2_Pos_M - 5.0) <= 15.0, 'residu 14,25 m -> aucun depassement de butee');

    (* --- Residu 14,75 m (haut de bande fermee) --- *)
    M2_Pos_M := 14.75 + 5.0;
    FOR i := 1 TO 800 DO
        FB_Bench(Enable := TRUE, RawPosM1 := RawPosM1, RawPosM2 := RawPosM2,
                 M1_RelayFwd := TRUE, M2_RelayFwd := TRUE,
                 M1_BrakeCmd := TRUE, M2_BrakeCmd := TRUE,
                 SimWinchCouplingModelActive := TRUE,
                 M1_CablePos_M := 5.0, M2_CablePos_M := M2_Pos_M,
                 BucketOffsetCloseM := 15.0, BucketCoherenceLimitM := 1.0);
        ASSERT_TRUE(FB_Bench.WinchCouplingCorrectionPts <= 82, 'correction bornee a 0,02 m par scan');
        M2_Pos_M := M2_Pos_M + DINT_TO_REAL(FB_Bench.WinchCouplingCorrectionPts) * (2.0 / 8192.0);
    END_FOR;
    ADVANCE_TIME(10000000);
    ASSERT_TRUE((M2_Pos_M - 5.0) >= 14.97, 'residu 14,75 m -> butee atteinte (ecart <= 0,2 %)');
    ASSERT_TRUE((M2_Pos_M - 5.0) <= 15.0, 'residu 14,75 m -> aucun depassement de butee');
END_TEST

TEST 'TC-P13-076 T419 ouverture M2 seule : roulis couvre l anticipation benne configuree'
VAR
    i                    : INT;
    RawPosAfterCommand   : UDINT;
    CoastDistanceActual_M : REAL;
END_VAR
    (* Un scan de descente relative charge la distance de roulis configuree dans
       FB_Sim_Encoder ; apres coupure, le codeur doit parcourir cette distance. *)
    RawPosM1 := 10000000;
    RawPosM2 := 50000000;
    FB_Bench(Enable := TRUE, RawPosM1 := RawPosM1, RawPosM2 := RawPosM2,
             M2_RelayFwd := FALSE, M2_RelayRev := TRUE, M2_StepNumber := 1,
             SimWinchCouplingModelActive := TRUE,
             SimWinchCoast_M := 0.35,
             M1_CablePos_M := 5.0, M2_CablePos_M := 6.31,
             BucketOffsetOpen_M := 0.0, BucketOpenAnticipation_M := 1.3,
             BucketAx15bOpenActive := TRUE);
    ASSERT_NEAR(FB_Bench.M2EffectiveCoastDistance_M, 1.3, 0.001,
                'fin AX15B -> roulis compense le scan mesure en retard');
    RawPosAfterCommand := RawPosM2;
    ADVANCE_TIME(10000000);

    FOR i := 1 TO 160 DO
        FB_Bench(Enable := TRUE, RawPosM1 := RawPosM1, RawPosM2 := RawPosM2,
                 M2_RelayFwd := FALSE, M2_RelayRev := FALSE, M2_StepNumber := 0,
                 SimWinchCouplingModelActive := TRUE,
                 SimWinchCoast_M := 0.35,
                 M1_CablePos_M := 5.0, M2_CablePos_M := 6.3,
                 BucketOffsetOpen_M := 0.0, BucketOpenAnticipation_M := 1.3,
                 BucketAx15bOpenActive := FALSE);
        ADVANCE_TIME(10000000);
    END_FOR;
    CoastDistanceActual_M := DINT_TO_REAL(UDINT_TO_DINT(RawPosAfterCommand)
                                          - UDINT_TO_DINT(RawPosM2)) * (2.0 / 8192.0);
    ASSERT_NEAR(CoastDistanceActual_M, 1.3, 0.03,
                'distance parcourue apres coupure atteint la butee ouverte');

    (* Un mouvement unitaire M2 hors demande auto garde son roulis de base. *)
    FB_Bench(Enable := TRUE, RawPosM1 := RawPosM1, RawPosM2 := RawPosM2,
             M2_RelayFwd := FALSE, M2_RelayRev := TRUE, M2_StepNumber := 1,
             SimWinchCouplingModelActive := TRUE,
             SimWinchCoast_M := 0.35,
             M1_CablePos_M := 5.0, M2_CablePos_M := 6.31,
             BucketOffsetOpen_M := 0.0, BucketOpenAnticipation_M := 1.3,
             BucketAx15bOpenActive := FALSE);
    ASSERT_NEAR(FB_Bench.M2EffectiveCoastDistance_M, FB_Bench.M2_EffectiveCoastM, 0.001,
                'jog manuel M2 -> roulis de base conserve');
END_TEST

(* ---- test_fb_simbench_m3_dynamics.st ---- *)
(* T417 — scénario d'intégration M3 isolé du test M2 historique.
   Il rejoue la chronologie de commande établie dans le code source :
   arrêt de demande avec frein maintenu desserré, puis demande de serrage.
   Pente nulle : ce test ne calibre ni ne reproduit un déplacement terrain. *)
SETUP
VAR
    FB_Bench : FB_SimBench;
    RawPosM1 : UDINT := 0;
    RawPosM2 : UDINT := 0;
END_VAR
END_SETUP

TEST 'T417-INT-010 M3 : rampe puis frein mecanique suivant la chronologie AX14-AX15'
VAR
    i : INT;
    PositionAfterStop_M : REAL;
END_VAR
    (* Repli deterministe P1, puis marche M3 : la DI frein ne doit pas anticiper. *)
    FB_Bench(Enable := FALSE, RawPosM1 := RawPosM1, RawPosM2 := RawPosM2);
    FOR i := 1 TO 30 DO
        FB_Bench(Enable := TRUE, M3_ReqTremie := TRUE, M3_ReqMaintenance := FALSE,
                 M3_SpeedCmd_Pct := 20.0, M3_BrakeCmd := TRUE,
                 SimM3SpeedFactor := 1.0, SimM3Slope_Mps2 := 0.0,
                 RawPosM1 := RawPosM1, RawPosM2 := RawPosM2);
    END_FOR;
    ASSERT_TRUE(FB_Bench.Translation.M3_BrakeIsOpen_DI,
                'Commande de desserrage maintenue : le contact frein finit ouvert');
    ASSERT_EQ(FB_Bench.Translation.M3_StatusWord, 16#0087,
              'La frequence active publie le status de marche');

    (* AX14 annule la demande ; avant AX15, la commande frein reste desserree. *)
    FOR i := 1 TO 80 DO
        FB_Bench(Enable := TRUE, M3_ReqTremie := FALSE, M3_ReqMaintenance := FALSE,
                 M3_SpeedCmd_Pct := 0.0, M3_BrakeCmd := TRUE,
                 SimM3SpeedFactor := 1.0, SimM3Slope_Mps2 := 0.0,
                 RawPosM1 := RawPosM1, RawPosM2 := RawPosM2);
    END_FOR;
    ASSERT_EQ(FB_Bench.Translation.M3_StatusWord, 16#0080,
              'La rampe a atteint l arret avant la fermeture mecanique');
    ASSERT_TRUE(FB_Bench.Translation.M3_BrakeIsOpen_DI,
                'Le frein reste ouvert tant que l automate le commande desserre');
    PositionAfterStop_M := FB_Bench.M3ObsPositionTrue_M;

    (* AX15 retire le desserrage : le contact ne peut pas retomber au premier scan. *)
    FB_Bench(Enable := TRUE, M3_ReqTremie := FALSE, M3_ReqMaintenance := FALSE,
             M3_SpeedCmd_Pct := 0.0, M3_BrakeCmd := FALSE,
             SimM3SpeedFactor := 1.0, SimM3Slope_Mps2 := 0.0,
             RawPosM1 := RawPosM1, RawPosM2 := RawPosM2);
    ASSERT_TRUE(FB_Bench.Translation.M3_BrakeIsOpen_DI,
                'Le delai mecanique interdit une fermeture du contact au premier scan');
    FOR i := 1 TO 20 DO
        FB_Bench(Enable := TRUE, M3_ReqTremie := FALSE, M3_ReqMaintenance := FALSE,
                 M3_SpeedCmd_Pct := 0.0, M3_BrakeCmd := FALSE,
                 SimM3SpeedFactor := 1.0, SimM3Slope_Mps2 := 0.0,
                 RawPosM1 := RawPosM1, RawPosM2 := RawPosM2);
    END_FOR;
    ASSERT_FALSE(FB_Bench.Translation.M3_BrakeIsOpen_DI,
                 'Apres le delai mecanique, le contact frein publie ferme');
    ASSERT_EQ(FB_Bench.M3ObsPositionTrue_M, PositionAfterStop_M,
              'Pente nulle : aucune derive inventee apres l arret variateur');
END_TEST
